Fanuc KAREL source: ka00118.KL

-- PROVISIONAL review KL for V770-1; original PC SHA256 9b1c1d22acccc1480cc60a8ad9be2940fefa82ec5eaefbdff19fffb432333e69
-- Incomplete behavior may be omitted. Consult companion uncertainty JSON. Do not deploy.
PROGRAM KA00118
%NOLOCKGROUP
-- UNRESOLVED_DECL SRC type=00001c
-- UNRESOLVED_DECL DST type=00001c
BEGIN
  -- UNRESOLVED_PC offsets 5-15; opcodes 9D,22,A5
  -- UNRESOLVED_PC offsets 20-32; opcodes 21,23
  -- UNRESOLVED_PC offsets 37-41; opcodes 7F
END KA00118
